(* IEC 61131-3 sources: Versio-VersionControlSystem/fixtures/projects/RefrigeratorControl/Device/Plc Logic/Application/Library/Alarm/DUTs, 4 files *)

(* ---- E_AlarmCategory.st ---- *)
{attribute 'qualified_only'}
{attribute 'strict'}
{attribute 'to_string'}
TYPE E_AlarmCategory :
(
	General 	:= 0,
	Power 		:= 1,
	Safety 		:= 2,
	Comms 		:= 3,
	Hardware 	:= 4
);
END_TYPE

(* ---- E_AlarmSeverity.st ---- *)
{attribute 'qualified_only'}
{attribute 'strict'}
{attribute 'to_string'}
TYPE E_AlarmSeverity :
(
	Diagnostic	 	:= 1,
	Low				:= 2,
	Medium			:= 3,
	High			:= 4
);
END_TYPE

(* ---- E_AlarmState.st ---- *)
{attribute 'qualified_only'}
{attribute 'strict'}
{attribute 'to_string'}
TYPE E_AlarmState :
(
	Off 		:= 0,
	Active 		:= 1
);
END_TYPE

(* ---- ST_AlarmSettings.st ---- *)
TYPE ST_AlarmSettings :
STRUCT
	ShortDesc			: STRING(20);
	Severity			: E_AlarmSeverity;
	Category			: E_AlarmCategory;
	Latch				: BOOL := FALSE;
	OnDelayTime			: TIME := T#0S;
	OffDelayTime		: TIME := T#0S;
	Enable				: BOOL := TRUE;
END_STRUCT
END_TYPE
